// TIA Portal V20 export
VAR_GLOBAL   // PLC tag table "COGNEX_FOLIE_P"
   "COG_FOLIE_P_COG_FOLIE_P_is3800-TriggerEnable" AT %Q10.0 : Bool;
   "COG_FOLIE_P_is3800-Trigger" AT %Q10.1 : Bool;
   "COG_FOLIE_P_is3800-ClearExposureComplete" AT %Q10.2 : Bool;
   "COG_FOLIE_P_is3800-Set Offline" AT %Q10.7 : Bool;
   "COG_FOLIE_P_is3800-TriggerReady" AT %I22.0 : Bool;
   "COG_FOLIE_P_is3800-TriggerAck" AT %I22.1 : Bool;
   "COG_FOLIE_P_is3800-ExposureComplete" AT %I22.2 : Bool;
   "COG_FOLIE_P_is3800-AcquCOG_FOLIE_P_isitionError" AT %I22.3 : Bool;
   "COG_FOLIE_P_is3800-Offline Reason" AT %I22.4 : Bool;
   "COG_FOLIE_P_is3800-Offline Reason(1)" AT %I22.5 : Bool;
   "COG_FOLIE_P_is3800-Offline Reason(2)" AT %I22.6 : Bool;
   "COG_FOLIE_P_is3800-Online" AT %I22.7 : Bool;
   "COG_FOLIE_P_is3800-AcquCOG_FOLIE_P_isitionID" AT %IW24 : Int;
   "COG_FOLIE_P_is3800-BufferResultsEnable" AT %Q11.0 : Bool;
   "COG_FOLIE_P_is3800-InspectionResultsAck" AT %Q11.1 : Bool;
   "COG_FOLIE_P_is3800-SetUserData" AT %Q11.2 : Bool;
   "COG_FOLIE_P_is3800-ExecuteCommand/JobLoad" AT %Q11.3 : Bool;
   "COG_FOLIE_P_is3800-ClearError" AT %Q11.7 : Bool;
   "COG_FOLIE_P_is3800-Reserved" AT %I26.0 : Bool;
   "COG_FOLIE_P_is3800-InspectionCompleted" AT %I26.1 : Bool;
   "COG_FOLIE_P_is3800-ResultsBufferOverrun" AT %I26.2 : Bool;
   "COG_FOLIE_P_is3800-ResultsValid" AT %I26.3 : Bool;
   "COG_FOLIE_P_is3800-CommandExecuting" AT %I26.4 : Bool;
   "COG_FOLIE_P_is3800-CommandCompleted" AT %I26.5 : Bool;
   "COG_FOLIE_P_is3800-CommandFailed" AT %I26.6 : Bool;
   "COG_FOLIE_P_is3800-SetUserDataAck" AT %I26.7 : Bool;
   "COG_FOLIE_P_is3800-ResultsPassed (Job)" AT %I27.0 : Bool;
   "COG_FOLIE_P_is3800-SystemValidated" AT %I27.1 : Bool;
   "COG_FOLIE_P_is3800-Error" AT %I27.7 : Bool;
   "COG_FOLIE_P_is3800-ErrorCode" AT %IW28 : Word;
   "COG_FOLIE_P_is3800-CommandID" AT %QW196 : Word;
   "COG_FOLIE_P_is3800-Current Job ID" AT %IW212 : Word;
   "COG_FOLIE_P_is3800-CommandResultCode" AT %IW214 : Word;
   "COG_FOLIE_P_is3800-ExternalEvent[0]" AT %Q12.0 : Bool;
   "COG_FOLIE_P_is3800-ExternalEvent[1]" AT %Q12.1 : Bool;
   "COG_FOLIE_P_is3800-ExternalEvent[2]" AT %Q12.2 : Bool;
   "COG_FOLIE_P_is3800-ExternalEvent[3]" AT %Q12.3 : Bool;
   "COG_FOLIE_P_is3800-ExternalEvent[4]" AT %Q12.4 : Bool;
   "COG_FOLIE_P_is3800-ExternalEvent[5]" AT %Q12.5 : Bool;
   "COG_FOLIE_P_is3800-ExternalEvent[6]" AT %Q12.6 : Bool;
   "COG_FOLIE_P_is3800-ExternalEvent[7]" AT %Q12.7 : Bool;
   "COG_FOLIE_P_is3800-ExternalEventAck[0]" AT %I30.0 : Bool;
   "COG_FOLIE_P_is3800-ExternalEventAck[1]" AT %I30.1 : Bool;
   "COG_FOLIE_P_is3800-ExternalEventAck[2]" AT %I30.2 : Bool;
   "COG_FOLIE_P_is3800-ExternalEventAck[3]" AT %I30.3 : Bool;
   "COG_FOLIE_P_is3800-ExternalEventAck[4]" AT %I30.4 : Bool;
   "COG_FOLIE_P_is3800-ExternalEventAck[5]" AT %I30.5 : Bool;
   "COG_FOLIE_P_is3800-ExternalEventAck[6]" AT %I30.6 : Bool;
   "COG_FOLIE_P_is3800-ExternalEventAck[7]" AT %I30.7 : Bool;
   "COG_FOLIE_P_is3800-UserData[0]" AT %QB198 : Byte;
   "COG_FOLIE_P_is3800-UserData[1]" AT %QB199 : Byte;
   "COG_FOLIE_P_is3800-UserData[2]" AT %QB200 : Byte;
   "COG_FOLIE_P_is3800-UserData[3]" AT %QB201 : Byte;
   "COG_FOLIE_P_is3800-UserData[4]" AT %QB202 : Byte;
   "COG_FOLIE_P_is3800-UserData[5]" AT %QB203 : Byte;
   "COG_FOLIE_P_is3800-UserData[6]" AT %QB204 : Byte;
   "COG_FOLIE_P_is3800-UserData[7]" AT %QB205 : Byte;
   "COG_FOLIE_P_is3800-UserData[8]" AT %QB206 : Byte;
   "COG_FOLIE_P_is3800-UserData[9]" AT %QB207 : Byte;
   "COG_FOLIE_P_is3800-UserData[10]" AT %QB208 : Byte;
   "COG_FOLIE_P_is3800-UserData[11]" AT %QB209 : Byte;
   "COG_FOLIE_P_is3800-UserData[12]" AT %QB210 : Byte;
   "COG_FOLIE_P_is3800-UserData[13]" AT %QB211 : Byte;
   "COG_FOLIE_P_is3800-UserData[14]" AT %QB212 : Byte;
   "COG_FOLIE_P_is3800-UserData[15]" AT %QB213 : Byte;
   "COG_FOLIE_P_is3800-InspectionID" AT %IW216 : Word;
   "COG_FOLIE_P_is3800-InspectionResultsCode" AT %IW218 : Int;
   "COG_FOLIE_P_is3800-InspectionResults[0]" AT %IB220 : Byte;
   "COG_FOLIE_P_is3800-InspectionResults[1]" AT %IB221 : Byte;
   "COG_FOLIE_P_is3800-InspectionResults[2]" AT %IB222 : Byte;
   "COG_FOLIE_P_is3800-InspectionResults[3]" AT %IB223 : Byte;
   "COG_FOLIE_P_is3800-InspectionResults[4]" AT %IB224 : Byte;
   "COG_FOLIE_P_is3800-InspectionResults[5]" AT %IB225 : Byte;
   "COG_FOLIE_P_is3800-InspectionResults[6]" AT %IB226 : Byte;
   "COG_FOLIE_P_is3800-InspectionResults[7]" AT %IB227 : Byte;
   "COG_FOLIE_P_is3800-InspectionResults[8]" AT %IB228 : Byte;
   "COG_FOLIE_P_is3800-InspectionResults[9]" AT %IB229 : Byte;
   "COG_FOLIE_P_is3800-InspectionResults[10]" AT %IB230 : Byte;
   "COG_FOLIE_P_is3800-InspectionResults[11]" AT %IB231 : Byte;
   "COG_FOLIE_P_is3800-InspectionResults[12]" AT %IB232 : Byte;
   "COG_FOLIE_P_is3800-InspectionResults[13]" AT %IB233 : Byte;
   "COG_FOLIE_P_is3800-InspectionResults[14]" AT %IB234 : Byte;
   "COG_FOLIE_P_is3800-InspectionResults[15]" AT %IB235 : Byte;
END_VAR
